// TIA Portal V21 export
// export: Created 2026-10-12T12:46:15.5115781Z, ExportSetting WithDefaults, DisplayName Totally Integrated Automation Portal, DisplayVersion V21, DisplayName STEP 7 Professional, DisplayVersion V21, DisplayName STEP 7 Safety, DisplayVersion V21, DisplayName Tech WebApplication, DisplayVersion V21, DisplayName WinCC Basic/Comfort/Advanced, DisplayVersion V21, DisplayName WinCC Unified, DisplayVersion V21
Screen "MANUAL"  800x480, Number=2, Template=MAIN
  ScreenLayer 
    Button "Button_1" at 166,194 size 179x82  Mode=Text, TextOff="CONVEYOR FWD JOG", TextOn="Text"
      RangeAppearanceAnimation "RangeAppearanceAnimation"
        tag DB_HMI_MOTOR JOG FWD PB
        1..1: back #00ff00, fore #000000
      on Press: SetBitWhileKeyPressed(Tag := DB_HMI_MOTOR JOG FWD PB, Bit := 0)
    Button "Button_2" at 429,190 size 179x82  Mode=Text, TextOff="CONVEYOR REV JOG", TextOn="Text"
      RangeAppearanceAnimation "RangeAppearanceAnimation"
        tag DB_HMI_MOTOR JOG REV PB
        1..1: back #00ff00, fore #000000
      on Press: SetBitWhileKeyPressed(Tag := DB_HMI_MOTOR JOG REV PB, Bit := 0)
    TextField "Template_Text field_2" at 308,62 size 210x27  Text="MANUAL OPERATION"
